// TIA Portal V20 export
Screen "190FX1Layout_Lifter"  1276x673
  ScreenItem "Line_Header_X0_Y64" at 0,64 size 1276x0  Type=HmiLine
  ScreenItem "permanentareaborderrectangle" at 0,0 size 0x0  Type=HmiRectangle
  ScreenItem "Button_Back" at 2,2 size 90x60  Type=HmiButton
  ScreenItem "Move_Legend" at 1183,2 size 90x60  Type=HmiButton
  ScreenItem "Fusszeile_Button_ManualOPMode1_2" at 188,2 size 90x60  Type=HmiButton
  ScreenItem "Fusszeile_Button_ManualOPMode1_1" at 95,2 size 90x60  Type=HmiButton
  ScreenItem "文本域_8" at 1172,-248 size 100x20  Type=HmiTextBox
  ScreenItem "文本域_9" at 1741,-563 size 100x20  Type=HmiTextBox
  ScreenItem "文本域_10" at 2310,-878 size 100x20  Type=HmiTextBox
  ScreenItem "文本域_12" at 321,1215 size 100x20  Type=HmiTextBox
  ScreenItem "Title_ScreenOverview_X390_Y2_1" at 384,2 size 510x57  Type=HmiTextBox
  ScreenItem "文本域_4" at 747,186 size 140x40  Type=HmiTextBox
  ScreenItem "文本域_6" at 747,451 size 140x40  Type=HmiTextBox
  ScreenItem "文本域_2" at 32,186 size 140x40  Type=HmiTextBox
  ScreenItem "文本域_3" at 32,451 size 140x40  Type=HmiTextBox
  ScreenItem "Graphic view_1" at 194,171 size 287x375  Type=HmiGraphicView
  ScreenItem "Line_6" at 177,219 size 125x77  Type=HmiLine
  ScreenItem "Line_7" at 175,478 size 134x5  Type=HmiLine
  ScreenItem "Graphic view_2" at 898,171 size 267x375  Type=HmiGraphicView
  ScreenItem "Line_1" at 887,383 size 115x90  Type=HmiLine
  ScreenItem "Line_2" at 887,207 size 109x157  Type=HmiLine
  ScreenItem "面板容器_1" at 35,228 size 142x51  Type=HmiFaceplateContainer
  ScreenItem "面板容器_3" at 35,493 size 142x51  Type=HmiFaceplateContainer
  ScreenItem "面板容器_4" at 747,230 size 142x51  Type=HmiFaceplateContainer
  ScreenItem "面板容器_5" at 747,493 size 142x51  Type=HmiFaceplateContainer
  ScreenItem "文本域_27" at -1,126 size 120x40  Type=HmiTextBox
  ScreenItem "文本域_5" at -1,82 size 120x40  Type=HmiTextBox
  ScreenItem "Button_Back_1" at 1180,606 size 90x60  Type=HmiButton
  ScreenItem "面板容器_2" at 1090,4 size 88x58  Type=HmiFaceplateContainer
  ScreenItem "OPMode1_Blocked" at 1164,6 size 14x14  Type=HmiGraphicView
  ScreenItem "OPMode4_Foreground_Blocked" at 1089,2 size 88x58  Type=HmiGraphicView
  ScreenItem "Fusszeile_Button_ManualOPMode1_3" at 987,1 size 90x60  Type=HmiButton
